Fanuc KAREL source: kc00036.KL

-- PROVISIONAL review KL for V770-1; original PC SHA256 768f8f5e6b9343969549af7ba94ea08286ecf87325733e51b06eeb52decd6af2
-- Incomplete behavior may be omitted. Consult companion uncertainty JSON. Do not deploy.
PROGRAM KC00036
%NOLOCKGROUP
BEGIN
  -- UNRESOLVED_PC offsets 5-15; opcodes 27,31,23
  -- UNRESOLVED_PC offsets 20-24; opcodes 7F
END KC00036
